// TIA Portal project "DEVOIR_TIA_PORTAL2" (V16)

(* hardware
DEVICE "Station S71500/ET200MP_1"  S7-1500 station
   slot 0: "Châssis_0"  Rack  6ES7 590-1***0-0AA0
   slot 1: "PLC_1"  CPU 1511C-1 PN  6ES7 511-1CK00-0AB0  V2.8
      slot 3: "Ecran CPU_1"  6ES7591-1AA00-0AA0
      slot 32768: "Interface PROFINET_1"  X1
         slot 32769: "Port_1"  X1 P1
         slot 32770: "Port_2"  X1 P2
      slot 34817: "Virtual CP interface port_1"  Virtual CP interface port  Virtual CP interface port
*)

// ===== PLC "PLC_1"  CPU 1511C-1 PN =====

VAR_GLOBAL   // PLC tag table "Table de variables standard"
   "S1" AT %I10.1 : Bool;
   "KM1" AT %Q4.1 : Bool;
   "KM2" AT %Q4.2 : Bool;
   "H1" AT %Q4.3 : Bool;
   "H2" AT %Q4.4 : Bool;
   "H3" AT %Q4.5 : Bool;
   "Tag_1" AT %M0.1 : Bool;
END_VAR

DATA_BLOCK "GRAFCET_DB"   // DB2
{ S7_Optimized_Access := 'TRUE' }
VERSION : 0.1
// stored: InstanceOfName GRAFCET
"GRAFCET"
BEGIN
END_DATA_BLOCK

// folder: System blocks/Program resources

DATA_BLOCK "C1"   // DB1
{ S7_Optimized_Access := 'TRUE' }
AUTHOR : Simatic
FAMILY : IEC
NAME : CNTR
VERSION : 1.0
// stored: InstanceOfName IEC_COUNTER
"IEC_COUNTER"
BEGIN
END_DATA_BLOCK

// folder: (top level)

FUNCTION_BLOCK "GRAFCET"   // FB1, GRAPH_PLUS
{ S7_Optimized_Access := 'TRUE' }
VERSION : 0.1
   VAR_INPUT
      OFF_SQ : Bool := false;   // Désactiver le graphe
      INIT_SQ : Bool := false;   // Mettre le graphe à l'état initial
      ACK_EF : Bool := false;   // Acquitter toutes les erreurs et perturbations
      S_PREV : Bool := false;   // Afficher l'étape précédente dans le paramètre S_NO
      S_NEXT : Bool := false;   // Afficher l'étape suivante dans le paramètre S_NO
      SW_AUTO : Bool := false;   // Mode automatique
      SW_TAP : Bool := false;   // Mode semi-automatique/Activation de l'étape suivante avec transition
      SW_TOP : Bool := false;   // Mode semi-automatique/Ignorer la transition
      SW_MAN : Bool := false;   // Mode manuel
      S_SEL : Int := 0;   // Sélectionner l'étape à afficher dans S_NO
      S_ON : Bool := false;   // Activer l'étape figurant dans le paramètre S_NO
      S_OFF : Bool := false;   // Désactiver l'étape figurant dans le paramètre S_NO
      T_PUSH : Bool := false;   // Validation de commutation pour transition en mode semi-automatique
   END_VAR
   VAR_OUTPUT
      S_NO : Int := 0;   // Numéro d'étape
      S_MORE : Bool := false;   // Il existe d'autres étapes qui peuvent être affichées dans S_NO.
      S_ACTIVE : Bool := false;   // L'étape affichée dans le paramètre S_NO est activée
      ERR_FLT : Bool := false;   // Erreur groupée Interlock or Supervision
      AUTO_ON : Bool := false;   // Mode automatique activé
      TAP_ON : Bool := false;   // Mode semi-automatique/Etape avec transition activé
      TOP_ON : Bool := false;   // Mode semi-automatique/Ignorer la transition activé
      MAN_ON : Bool := false;   // Mode manuel activé
   END_VAR
   VAR
      HMI_INFO : Array[0..0] of UInt;
      RT_DATA : G7_RTDataPlus_V6;   // Plage de données interne
      Trans1 : G7_TransitionPlus_V6;   // Structure de la transition
      step1 : G7_StepPlus_V6;   // Structure de l'étape
      Step2 : G7_StepPlus_V6;   // Structure de l'étape
      Trans2 : G7_TransitionPlus_V6;   // Structure de la transition
      Step3 : G7_StepPlus_V6;   // Structure de l'étape
      Trans3 : G7_TransitionPlus_V6;   // Structure de la transition
      Step20 : G7_StepPlus_V6;   // Structure de l'étape
      Step10 : G7_StepPlus_V6;   // Structure de l'étape
      Trans4 : G7_TransitionPlus_V6;   // Structure de la transition
      Step11 : G7_StepPlus_V6;   // Structure de l'étape
      Trans5 : G7_TransitionPlus_V6;   // Structure de la transition
      Step12 : G7_StepPlus_V6;   // Structure de l'étape
      Trans7 : G7_TransitionPlus_V6;   // Structure de la transition
      Step21 : G7_StepPlus_V6;   // Structure de l'étape
      Trans8 : G7_TransitionPlus_V6;   // Structure de la transition
      Step22 : G7_StepPlus_V6;   // Structure de l'étape
      Trans10 : G7_TransitionPlus_V6;   // Structure de la transition
      Step4 : G7_StepPlus_V6;   // Structure de l'étape
      Trans11 : G7_TransitionPlus_V6;   // Structure de la transition
      Trans12 : G7_TransitionPlus_V6;   // Structure de la transition
      Trans9 : G7_TransitionPlus_V6;   // Structure de la transition
   END_VAR
BEGIN
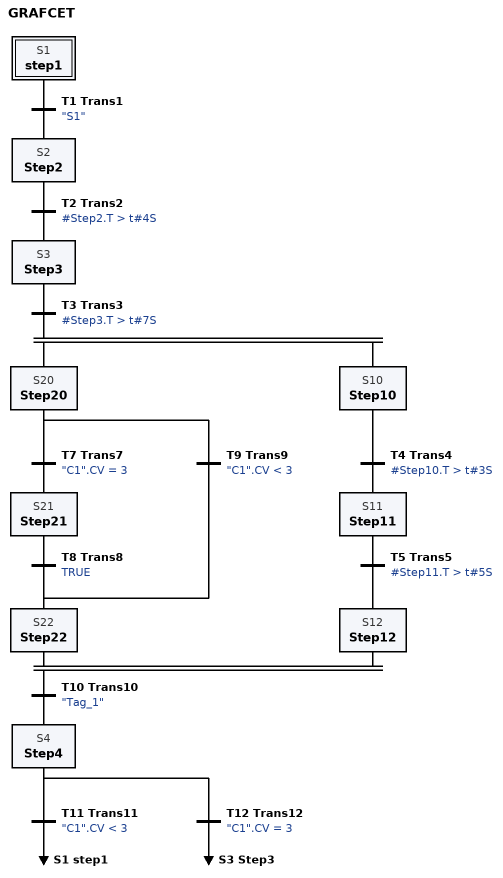
   // sequencer 1
   INITIAL_STEP step1:   // S1, max time T#10S, warning time T#7S
   END_STEP
   TRANSITION Trans1 FROM step1 TO Step2   // T1
      := "S1";
   END_TRANSITION
   STEP Step2:   // S2, max time T#10S, warning time T#7S
   END_STEP
   TRANSITION Trans2 FROM Step2 TO Step3   // T2
      := #Step2.T > t#4S;
   END_TRANSITION
   STEP Step3:   // S3, max time T#10S, warning time T#7S
   END_STEP
   TRANSITION Trans3 FROM Step3 TO (Step20, Step10)   // T3
      := #Step3.T > t#7S;
   END_TRANSITION
   STEP Step20:   // S20, max time T#10S, warning time T#7S
   END_STEP
   TRANSITION Trans7 FROM Step20 TO Step21   // T7
      := "C1".CV = 3;
   END_TRANSITION
   TRANSITION Trans9 FROM Step20 TO Step22   // T9
      := "C1".CV < 3;
   END_TRANSITION
   STEP Step10:   // S10, max time T#10S, warning time T#7S
   END_STEP
   TRANSITION Trans4 FROM Step10 TO Step11   // T4
      := #Step10.T > t#3S;
   END_TRANSITION
   STEP Step11:   // S11, max time T#10S, warning time T#7S
   END_STEP
   TRANSITION Trans5 FROM Step11 TO Step12   // T5
      := #Step11.T > t#5S;
   END_TRANSITION
   STEP Step12:   // S12, max time T#10S, warning time T#7S
   END_STEP
   STEP Step21:   // S21, max time T#10S, warning time T#7S
   END_STEP
   TRANSITION Trans8 FROM Step21 TO Step22   // T8
      := TRUE;
   END_TRANSITION
   STEP Step22:   // S22, max time T#10S, warning time T#7S
   END_STEP
   TRANSITION Trans10 FROM (Step12, Step22) TO Step4   // T10
      := "Tag_1";
   END_TRANSITION
   STEP Step4:   // S4, max time T#10S, warning time T#7S
   END_STEP
   TRANSITION Trans11 FROM Step4 TO step1   // T11, jump
      := "C1".CV < 3;
   END_TRANSITION
   TRANSITION Trans12 FROM Step4 TO Step3   // T12, jump
      := "C1".CV = 3;
   END_TRANSITION
END_FUNCTION_BLOCK

FUNCTION "COMPTEUR" : Void   // FC1, LAD
{ S7_Optimized_Access := 'TRUE' }
VERSION : 0.1
BEGIN

REGION Network 1
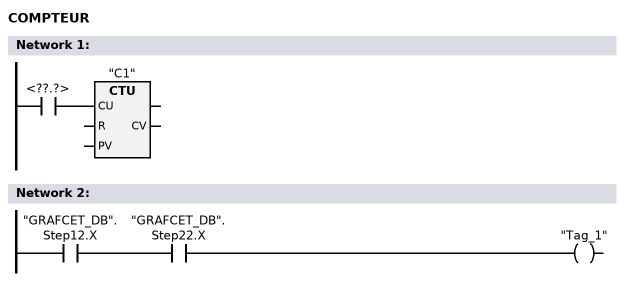
   // no checked SCL form for this network; see the picture
END_REGION

REGION Network 2
   RUNG wire#powerrail
      Contact( "GRAFCET_DB".Step12.X )
      Contact( "GRAFCET_DB".Step22.X )
      Coil( "Tag_1" )
   END_RUNG
   // the same network as SCL:
   "Tag_1" := "GRAFCET_DB".Step12.X AND "GRAFCET_DB".Step22.X;
END_REGION
END_FUNCTION

ORGANIZATION_BLOCK "Main"   // OB1, LAD, ProgramCycle
TITLE = "Main Program Sweep (Cycle)"
{ S7_Optimized_Access := 'TRUE' }
VERSION : 0.1
   VAR_INPUT
      Initial_Call : Bool;   // Initial call of this OB
      Remanence : Bool;   // =True, if remanent data are available
   END_VAR
BEGIN

REGION Network 1
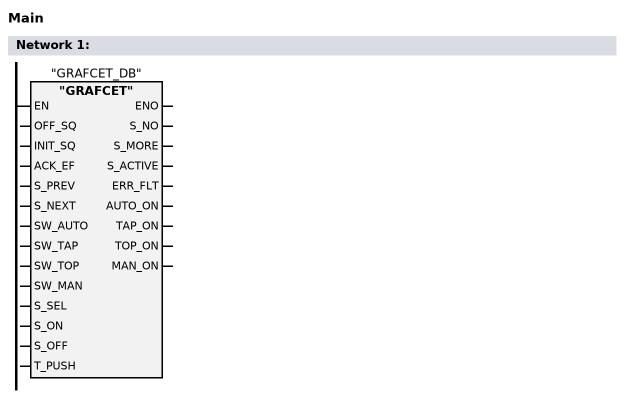
   RUNG wire#powerrail
      "GRAFCET_DB"(OFF_SQ :=, INIT_SQ :=, ACK_EF :=, S_PREV :=, S_NEXT :=, SW_AUTO :=, SW_TAP :=, SW_TOP :=, SW_MAN :=, S_SEL :=, S_ON :=, S_OFF :=, T_PUSH :=, S_NO =>, S_MORE =>, S_ACTIVE =>, ERR_FLT =>, AUTO_ON =>, TAP_ON =>, TOP_ON =>, MAN_ON =>)
   END_RUNG
   // the same network as SCL:
   "GRAFCET_DB"();   // "GRAFCET"
END_REGION
END_ORGANIZATION_BLOCK